// TIA Portal V20 export
// export: Created 2026-10-12T05:35:25.9325808Z, ExportSetting WithDefaults, DisplayName Totally Integrated Automation Portal, DisplayVersion V20, DisplayName TIA Portal Openness, DisplayVersion V20, DisplayName TIA Portal Teamcenter Gateway, DisplayVersion V20, DisplayName TIA Portal Version Control Interface, DisplayVersion V20, DisplayName SINAMICS Startdrive Advanced, DisplayVersion V20 SP1 Update 2, DisplayName SINAMICS Startdrive G110M, G120, G120C, G120D, G120P, G115D, DisplayVersion V20 SP1 Update 2, DisplayName SINAMICS Startdrive G130, G150, S120, S150, SINAMICS MV, G220, S200, S210, DisplayVersion V20 SP1 Update 2, DisplayName STEP 7 Professional, DisplayVersion V20, DisplayName STEP 7 Safety, DisplayVersion V20, DisplayName WinCC Basic/Comfort/Advanced, DisplayVersion V20, DisplayName WinCC Professional, DisplayVersion V20, DisplayName WinCC Unified, DisplayVersion V20
FUNCTION "FRK_JsonAdd" : Bool   // FC110, SCL
{ S7_Optimized_Access := 'TRUE' }
VERSION : 0.1
// stored: AutoNumber true, IsIECCheckEnabled false, SetENOAutomatically false, UDAEnableTagReadback false
   VAR_INPUT
      Key : String;
      Value : WString;
      Quoted : Bool;
      LastField : Bool;
   END_VAR
   VAR_IN_OUT
      Line : WString;
   END_VAR
   VAR_TEMP
      Index : Int;
      Ch : WChar;
      FirstChar : Int;
      Piece : WString[2];
      Ok : Bool;
   END_VAR
BEGIN

   #FRK_JsonAdd := FALSE;
   #Ok := "FRK_JsonPut"(Text := CONCAT(IN1 := WSTRING#'"', IN2 := STRING_TO_WSTRING(#Key), IN3 := WSTRING#'":'), Line := #Line);
   IF NOT #Ok THEN
       RETURN;
   END_IF;
   IF #Quoted THEN
       #Ok := "FRK_JsonPut"(Text := WSTRING#'"', Line := #Line);
       IF NOT #Ok THEN
           RETURN;
       END_IF;
   END_IF;
   #FirstChar := 1;
   // Siemens integer conversions include a leading '+'. JSON numbers do not.
   IF NOT #Quoted THEN
       IF LEN(#Value) = 0 THEN
           RETURN;
       END_IF;
       IF #Value[1] = WCHAR#'+' THEN
           #FirstChar := 2;
       END_IF;
       IF #FirstChar > LEN(#Value) THEN
           RETURN;
       END_IF;
   END_IF;
   FOR #Index := #FirstChar TO LEN(#Value) DO
       #Ch := #Value[#Index];
       #Piece := WSTRING#' ';
       #Piece[1] := #Ch;
       IF NOT #Quoted AND (#Ch < WCHAR#'0' OR #Ch > WCHAR#'9') THEN
           RETURN;
       END_IF;
       IF #Quoted THEN
           IF #Ch = WCHAR#'"' THEN
               #Piece := WSTRING#'\"';
           ELSIF #Ch = WCHAR#'\' THEN
               #Piece := WSTRING#'\\';
           ELSIF #Ch = WCHAR#'$000A' THEN
               #Piece := WSTRING#'\n';
           ELSIF #Ch = WCHAR#'$000D' THEN
               #Piece := WSTRING#'\r';
           ELSIF #Ch = WCHAR#'$0009' THEN
               #Piece := WSTRING#'\t';
           ELSIF #Ch = WCHAR#'$0008' THEN
               #Piece := WSTRING#'\b';
           ELSIF #Ch = WCHAR#'$000C' THEN
               #Piece := WSTRING#'\f';
           ELSIF #Ch < WCHAR#'$0020' THEN
               RETURN;
           END_IF;
       END_IF;
       #Ok := "FRK_JsonPut"(Text := #Piece, Line := #Line);
       IF NOT #Ok THEN
           RETURN;
       END_IF;
   END_FOR;
   IF #Quoted THEN
       #Ok := "FRK_JsonPut"(Text := WSTRING#'"', Line := #Line);
       IF NOT #Ok THEN
           RETURN;
       END_IF;
   END_IF;
   IF #LastField THEN
       #Piece := WSTRING#'}';
   ELSE
       #Piece := WSTRING#',';
   END_IF;
   #FRK_JsonAdd := "FRK_JsonPut"(Text := #Piece, Line := #Line);
END_FUNCTION
